FUNCTION_BLOCK FB_System_Time
VAR_OUTPUT
    Delta_Time : LREAL := 0;
	now : ULINT := 0;
END_VAR
VAR
    Last_Time : ULINT := 0;
	ConversionFactorSeconds : LREAL := 1E-7;
END_VAR

// FB must be called every PLC cycle, prefferably in the main() function.

now := Tc2_System.F_GetSystemTime();

IF Last_Time > 0 THEN
    Delta_Time := TO_LREAL(now - Last_Time) * ConversionFactorSeconds;
ELSE
    Delta_Time := 0;
END_IF

Last_Time := now;

END_FUNCTION_BLOCK

(* stored: Version 1.1.0.1, ProductVersion 3.1.4024.13
   POU FB_System_Time: Id {5538c938-e0ce-479c-836f-7e403d8ebc09}, SpecialFunc None *)
